// TIA Portal V20 export
FUNCTION "POS3_0_Betriebsart" : Void   // FC40, STL
{ S7_Optimized_Access := 'TRUE' }
BEGIN

NETWORK
TITLE = Schrittkette Halt von Betriebsart
      A(;
      A     "03_Betriebsart_DB".BA_Manuell;
      A(;
      L     "HMI_SYS"."Aktueller Bildschirm";
      L     21300;  // Bildschirm Einzelschritt ist aktiv
      ==I;
      );
      );

      O     "03_Betriebsart_DB".BA_Automatik;

      O(;  // Richten aktiv oder angefordert
      A     "03_Betriebsart_DB".BA_Richten;
      A(;
      A     "POS3_0_Signal".Station.SK_Richten_gestartet;
      O     "POS3_0_Signal".Station.SK_Freigabe_Richten;
      );
      );
      NOT;
      =     "POS3_0_Signal".Station.SK_Halt_von_Betriebsart;


NETWORK
TITLE = Schrittkettenaufruf
      ON    "03_Betriebsart_DB"."NOT-HALT OK";
      ON    "03_Betriebsart_DB"."Schutztüren OK";
      O     "03_Betriebsart_DB".BA_0;
      O     "POS3_0_Signal".Station.SK_Halt_von_Betriebsart;
      AN    "POS3_0_Signal".Schrittkette.SQ_HALTED;
      A     "Zyklisch wechselnder Merker";
      O(;
      A     "03_Betriebsart_DB"."NOT-HALT OK";
      A     "03_Betriebsart_DB"."Schutztüren OK";
      AN    "03_Betriebsart_DB".BA_0;
      AN    "POS3_0_Signal".Station.SK_Halt_von_Betriebsart;
      A     "POS3_0_Signal".Schrittkette.SQ_HALTED;
      A     "Zyklisch wechselnder Merker";
      );
      =     "POS3_0_Signal".Schrittkette.HALT_SQ;

      AN    "03_Betriebsart_DB"."NOT-HALT OK";
      ON    "03_Betriebsart_DB"."Schutztüren OK";
      O     "03_Betriebsart_DB".BA_0;
      O     "POS3_0_Signal".Station.SK_Halt_von_Betriebsart;
      AN    "POS3_0_Signal".Schrittkette.TM_HALTED;
      A     "Zyklisch wechselnder Merker";
      O(;
      A     "03_Betriebsart_DB"."NOT-HALT OK";
      A     "03_Betriebsart_DB"."Schutztüren OK";
      AN    "03_Betriebsart_DB".BA_0;
      AN    "POS3_0_Signal".Station.SK_Halt_von_Betriebsart;
      A     "POS3_0_Signal".Schrittkette.TM_HALTED;
      A     "Zyklisch wechselnder Merker";
      );
      =     "POS3_0_Signal".Schrittkette.HALT_TM;

      ON    "03_Betriebsart_DB"."NOT-HALT OK";
      ON    "03_Betriebsart_DB"."Schutztüren OK";
      O     "03_Betriebsart_DB".BA_0;
      O     "POS3_0_Signal".Station.SK_Halt_von_Betriebsart;
      AN    "POS3_0_Signal".Schrittkette.OP_ZEROED;
      A     "Zyklisch wechselnder Merker";
      O(;
      A     "03_Betriebsart_DB"."NOT-HALT OK";
      A     "03_Betriebsart_DB"."Schutztüren OK";
      AN    "03_Betriebsart_DB".BA_0;
      AN    "POS3_0_Signal".Station.SK_Halt_von_Betriebsart;
      A     "POS3_0_Signal".Schrittkette.OP_ZEROED;
      A     "Zyklisch wechselnder Merker";
      );
      =     "POS3_0_Signal".Schrittkette.ZERO_OP;





NETWORK
TITLE = Tipp/Autobetriebbetrieb
      A     "HMI_BETR_ART_POS".POS3_0.Taster_Anwahl_Tipp;
      AN    "POS3_0_Signal".Schrittkette.TAP_ON;
      A     "Zyklisch wechselnder Merker";
      =     "POS3_0_Signal".Schrittkette.SW_TAP;


      AN    "HMI_BETR_ART_POS".POS3_0.Taster_Anwahl_Tipp;
      AN    "POS3_0_Signal".Schrittkette.AUTO_ON;
      A     "Zyklisch wechselnder Merker";
      =     "POS3_0_Signal".Schrittkette.SW_AUTO;

NETWORK
TITLE = Tippen
      A     "03_Betriebsart_DB".Start_Taste_FP;
      O     "HMI_BETR_ART_POS".POS3_0.Taster_Tipp_Plus;
      =     "POS3_0_Signal".Schrittkette.T_PUSH;




NETWORK
TITLE = Tippen angewählt
END_FUNCTION
